(* IEC 61131-3 sources: 89152_FlorisHendrix_AfstudeerProject/89152_FlorisHendrix_ExamenProject/Stations/MachineControl/MachineControl/Drive, 2 files *)

(* ---- _DriveAxis1.st ---- *)
FUNCTION GLOBAL TAB DRIVETAB__DRIVEAXIS1
	1$UDINT, TO_UDINT(OFF(L1)-OFF(L0)),L0:
G01:	1$USINT,' '' '' '' ',
	2$USINT,' '' '' '' ',
	3$USINT,' '' '' '' ',
	4$USINT,1790$DINT,
	5$USINT,5400$DINT,
	6$USINT,6200$DINT,
	7$USINT,8$DINT,
	8$USINT,35$DINT,
	9$USINT,500$DINT,
	10$USINT,1500$DINT,
	11$USINT,24$DINT,
	13$USINT,2$DINT,
	14$USINT,177$DINT,
	15$USINT,1000$DINT,
	17$USINT,0$DINT,
	18$USINT,0$DINT,
	21$USINT,0$DINT,
	22$USINT,10$DINT,
	23$USINT,100$DINT,
G03:	32$USINT,3$DINT,
	33$USINT,50$DINT,
	35$USINT,18$DINT,
	36$USINT,75$DINT,
	38$USINT,108$DINT,
	41$USINT,65$DINT,
	42$USINT,10000$DINT,
	43$USINT,595582655$DINT,
	44$USINT,0$DINT,
	45$USINT,1073741824$DINT,
	46$USINT,67117056$DINT,
	47$USINT,300000$DINT,
	48$USINT,1$DINT,
	49$USINT,15$DINT,
	168$USINT,30$DINT,
	169$USINT,26$DINT,
	170$USINT,35$DINT,
G04:	50$USINT,5700$DINT,
	51$USINT,1400$DINT,
	53$USINT,70$DINT,
	56$USINT,1790$DINT,
	57$USINT,5400$DINT,
	59$USINT,85$DINT,
	167$USINT,100$DINT,
G05:	60$USINT,1000$DINT,
	61$USINT,1000$DINT,
	62$USINT,400$DINT,
	63$USINT,1000$DINT,
	64$USINT,80$DINT,
	65$USINT,4100$DINT,
	66$USINT,0$DINT,
	67$USINT,0$DINT,
	68$USINT,0$DINT,
G06:	70$USINT,10000$DINT,
	71$USINT,1005$DINT,
	72$USINT,16$DINT,
	73$USINT,1000$DINT,
	74$USINT,1000$DINT,
	75$USINT,3276800$DINT,
	76$USINT,0$DINT,
G08:	90$USINT,5000$DINT,
	91$USINT,775$DINT,
	92$USINT,0$DINT,
	93$USINT,3591$DINT,
	94$USINT,517$DINT,
	95$USINT,1000$DINT,
	99$USINT,100$DINT,
	103$USINT,2$DINT,
	105$USINT,600$DINT,
	108$USINT,' '' '' '' ',
	109$USINT,' '' '' '' ',
	110$USINT,' '' '' '' ',
	114$USINT,0$DINT,
	115$USINT,0$DINT,
	116$USINT,0$DINT,
	117$USINT,100$DINT,
	118$USINT,0$DINT,
	119$USINT,2500$DINT,
	120$USINT,300$DINT,
	121$USINT,2000$DINT,
	124$USINT,2386$DINT,
	164$USINT,0$DINT,
	165$USINT,0$DINT,
	173$USINT,0$DINT,
G14:	127$USINT,0$DINT,
	128$USINT,100$DINT,
	129$USINT,100$DINT,
	130$USINT,100$DINT,
	131$USINT,100$DINT,
	132$USINT,100$DINT,
	133$USINT,100$DINT,
	134$USINT,100$DINT,
	135$USINT,100$DINT,
	136$USINT,100$DINT,
	137$USINT,100$DINT,
	138$USINT,100$DINT,
	139$USINT,100$DINT,
	140$USINT,100$DINT,
	141$USINT,100$DINT,
	142$USINT,100$DINT,
	143$USINT,100$DINT,
	144$USINT,100$DINT,
	145$USINT,100$DINT,
	146$USINT,100$DINT,
	147$USINT,100$DINT,
	148$USINT,100$DINT,
	149$USINT,100$DINT,
	150$USINT,100$DINT,
	151$USINT,100$DINT,
	152$USINT,100$DINT,
	153$USINT,100$DINT,
	154$USINT,100$DINT,
	155$USINT,100$DINT,
	156$USINT,100$DINT,
	157$USINT,100$DINT,
	158$USINT,100$DINT,
	159$USINT,100$DINT,L1:
TO_UDINT(OFF(L3)-OFF(L2)),L2:
	01$USINT, OFF(G01),
	03$USINT, OFF(G03),
	04$USINT, OFF(G04),
	05$USINT, OFF(G05),
	06$USINT, OFF(G06),
	08$USINT, OFF(G08),
	14$USINT, OFF(G14),L3:
END_FUNCTION

(* ---- _DriveAxis2.st ---- *)
FUNCTION GLOBAL TAB DRIVETAB__DRIVEAXIS2
	1$UDINT, TO_UDINT(OFF(L1)-OFF(L0)),L0:
G01:	1$USINT,' '' '' '' ',
	2$USINT,' '' '' '' ',
	3$USINT,' '' '' '' ',
	4$USINT,1790$DINT,
	5$USINT,5400$DINT,
	6$USINT,6200$DINT,
	7$USINT,8$DINT,
	8$USINT,35$DINT,
	9$USINT,500$DINT,
	10$USINT,1500$DINT,
	11$USINT,24$DINT,
	13$USINT,2$DINT,
	14$USINT,93$DINT,
	15$USINT,1000$DINT,
	17$USINT,0$DINT,
	18$USINT,0$DINT,
	21$USINT,0$DINT,
	22$USINT,10$DINT,
	23$USINT,100$DINT,
G03:	32$USINT,3$DINT,
	33$USINT,50$DINT,
	35$USINT,18$DINT,
	36$USINT,0$DINT,
	38$USINT,85$DINT,
	41$USINT,65$DINT,
	42$USINT,10000$DINT,
	43$USINT,591388351$DINT,
	44$USINT,0$DINT,
	45$USINT,1073741824$DINT,
	46$USINT,71311360$DINT,
	47$USINT,3000000$DINT,
	48$USINT,1$DINT,
	49$USINT,0$DINT,
	168$USINT,60$DINT,
	169$USINT,55$DINT,
	170$USINT,55$DINT,
G04:	50$USINT,5700$DINT,
	51$USINT,1400$DINT,
	53$USINT,70$DINT,
	56$USINT,1790$DINT,
	57$USINT,5400$DINT,
	59$USINT,85$DINT,
	167$USINT,100$DINT,
G05:	60$USINT,14000$DINT,
	61$USINT,10000$DINT,
	62$USINT,400$DINT,
	63$USINT,1000$DINT,
	64$USINT,80$DINT,
	65$USINT,4100$DINT,
	66$USINT,0$DINT,
	67$USINT,0$DINT,
	68$USINT,0$DINT,
G06:	70$USINT,80000$DINT,
	71$USINT,1005$DINT,
	72$USINT,16$DINT,
	73$USINT,1000$DINT,
	74$USINT,1000$DINT,
	75$USINT,3276800$DINT,
	76$USINT,0$DINT,
G08:	90$USINT,5000$DINT,
	91$USINT,775$DINT,
	92$USINT,0$DINT,
	93$USINT,3591$DINT,
	94$USINT,517$DINT,
	95$USINT,1000$DINT,
	99$USINT,100$DINT,
	103$USINT,2$DINT,
	105$USINT,600$DINT,
	108$USINT,' '' '' '' ',
	109$USINT,' '' '' '' ',
	110$USINT,' '' '' '' ',
	114$USINT,0$DINT,
	115$USINT,0$DINT,
	116$USINT,0$DINT,
	117$USINT,100$DINT,
	118$USINT,0$DINT,
	119$USINT,2500$DINT,
	120$USINT,300$DINT,
	121$USINT,2000$DINT,
	124$USINT,0$DINT,
	164$USINT,0$DINT,
	165$USINT,0$DINT,
	173$USINT,0$DINT,
G14:	127$USINT,0$DINT,
	128$USINT,100$DINT,
	129$USINT,100$DINT,
	130$USINT,100$DINT,
	131$USINT,100$DINT,
	132$USINT,100$DINT,
	133$USINT,100$DINT,
	134$USINT,100$DINT,
	135$USINT,100$DINT,
	136$USINT,100$DINT,
	137$USINT,100$DINT,
	138$USINT,100$DINT,
	139$USINT,100$DINT,
	140$USINT,100$DINT,
	141$USINT,100$DINT,
	142$USINT,100$DINT,
	143$USINT,100$DINT,
	144$USINT,100$DINT,
	145$USINT,100$DINT,
	146$USINT,100$DINT,
	147$USINT,100$DINT,
	148$USINT,100$DINT,
	149$USINT,100$DINT,
	150$USINT,100$DINT,
	151$USINT,100$DINT,
	152$USINT,100$DINT,
	153$USINT,100$DINT,
	154$USINT,100$DINT,
	155$USINT,100$DINT,
	156$USINT,100$DINT,
	157$USINT,100$DINT,
	158$USINT,100$DINT,
	159$USINT,100$DINT,L1:
TO_UDINT(OFF(L3)-OFF(L2)),L2:
	01$USINT, OFF(G01),
	03$USINT, OFF(G03),
	04$USINT, OFF(G04),
	05$USINT, OFF(G05),
	06$USINT, OFF(G06),
	08$USINT, OFF(G08),
	14$USINT, OFF(G14),L3:
END_FUNCTION
